Fanuc KAREL source: ko00042.KL

-- PROVISIONAL review KL for V1013-1; original PC SHA256 d444eb81d94602734bf4c162ca9823197cf874c0f93f15c44f890b35503cc95c
-- Incomplete behavior may be omitted. Consult companion uncertainty JSON. Do not deploy.
PROGRAM KO00042
%NOLOCKGROUP
BEGIN
  -- UNRESOLVED_PC offsets 5-12; opcodes 9D,23
  -- UNRESOLVED_PC offsets 17-69; opcodes 27,27,49,7E,AD,27,49,7E,AD,22,31,7E,4A
  -- UNRESOLVED_PC offsets 74-78; opcodes 7F
END KO00042
